TYPE "ST_PressDemoOutImm"
VERSION : 0.1
   STRUCT
      Homed : Bool;
      TwoHandStartReady : Bool;
   END_STRUCT;

END_TYPE

